(*
SPDX-FileCopyrightText: © 2026 Oleksandr Tiutyk <trofimich@gmail.com>
SPDX-License-Identifier: MIT
License: https://opensource.org/license/mit
*)

(*!
<summary>
Beckhoff EL2502: 2-channel PWM output terminal (24 V DC, up to 20 kHz).
</summary>
<description>
Requires the duty-only Pulse width (standard) assignment, RxPDOs 0x1600 and 0x1601,
with signed presentation selected through CoE. Configure period/frequency before enabling outputs.
Cyclic-period and unsigned-presentation variants are outside this model.
When used for I/O, link located fields or their containing buffers to the matching selected PDOs.
The record is not a packed wire buffer; compiler padding is not part of the device specification.
Unlinked/default values do not prove valid I/O. The caller evaluates bus/channel validity before use.
Use one owner task per instance and externally synchronize other access; multi-field snapshots are not atomic.
Copies store data without creating hardware links. Keep borrowed field references valid while consumers are bound.
This passive record performs no validation, synchronization, configuration or protocol advancement.
</description>
*)
TYPE EL2502 :
STRUCT
	Ch1 : PWM_OUTPUT_CHANNEL;
	Ch2 : PWM_OUTPUT_CHANNEL;
END_STRUCT
END_TYPE

(* stored: Version 1.1.0.1, ProductVersion 3.1.4026.20
   DUT EL2502: Id {64b5244a-d4bb-4127-916b-7120a77cf490} *)
